// TIA Portal V20 export
Screen "OP02Pop-up_PRBHome"  274x350
  ScreenItem "Text field TG Status" at 1,0 size 273x47  Type=HmiTextBox
  ScreenItem "Cancel Mode" at 195,3 size 76x42  Type=HmiButton
  ScreenItem "Rectangle TG1" at 4,52 size 265x29  Type=HmiRectangle
  ScreenItem "Textfeld_1" at 9,57 size 21x20  Type=HmiTextBox
  ScreenItem "Textfeld_2" at 50,56 size 245x20  Type=HmiTextBox
  ScreenItem "Rectangle TG1_1" at 4,84 size 265x29  Type=HmiRectangle
  ScreenItem "Textfeld_5" at 9,89 size 21x20  Type=HmiTextBox
  ScreenItem "Rectangle TG1_2" at 4,116 size 265x29  Type=HmiRectangle
  ScreenItem "Textfeld_8" at 9,121 size 21x20  Type=HmiTextBox
  ScreenItem "Rectangle TG1_3" at 4,148 size 265x29  Type=HmiRectangle
  ScreenItem "Rectangle TG1_4" at 4,180 size 265x29  Type=HmiRectangle
  ScreenItem "Rectangle TG1_5" at 4,212 size 265x29  Type=HmiRectangle
  ScreenItem "Textfeld_18" at 10,153 size 21x20  Type=HmiTextBox
  ScreenItem "Textfeld_3" at 50,88 size 245x20  Type=HmiTextBox
  ScreenItem "Textfeld_4" at 50,121 size 245x20  Type=HmiTextBox
  ScreenItem "Textfeld_9" at 50,152 size 275x20  Type=HmiTextBox
  ScreenItem "Rectangle TG1_6" at 3,245 size 265x29  Type=HmiRectangle
  ScreenItem "Textfeld_6" at 10,185 size 21x20  Type=HmiTextBox
  ScreenItem "Textfeld_11" at 50,187 size 275x20  Type=HmiTextBox
  ScreenItem "Rectangle TG1_7" at 4,279 size 265x29  Type=HmiRectangle
  ScreenItem "Textfeld_10" at 10,217 size 21x20  Type=HmiTextBox
  ScreenItem "Textfeld_12" at 50,218 size 275x20  Type=HmiTextBox
  ScreenItem "Rectangle TG1_8" at 4,314 size 265x29  Type=HmiRectangle
  ScreenItem "Textfeld_16" at 10,250 size 21x20  Type=HmiTextBox
  ScreenItem "Textfeld_13" at 50,250 size 275x20  Type=HmiTextBox
  ScreenItem "Line_1" at 37,52 size 1x291  Type=HmiLine
